Fanuc KAREL source: kt00857.KL

-- PROVISIONAL review KL for V770-1; original PC SHA256 beacf136756bc76b702b1e8c7d108e6b8bc8b15ee67f3d41e52b0241ccb162a3
-- Incomplete behavior may be omitted. Consult companion uncertainty JSON. Do not deploy.
PROGRAM KT00857
%NOLOCKGROUP
VAR
  I1 : INTEGER
  I2 : INTEGER
  OUT : REAL
BEGIN
  -- UNRESOLVED_PC offsets 5-16; opcodes 2E,23
  -- UNRESOLVED_PC offsets 21-32; opcodes 2E,23
  -- UNRESOLVED_PC offsets 37-48; opcodes 2E,23
  -- UNRESOLVED_PC offsets 53-64; opcodes 2E,23
  -- UNRESOLVED_PC offsets 69-87; opcodes 27,27,21,64,76,64,23
  -- UNRESOLVED_PC offsets 92-96; opcodes 7F
END KT00857
